// TIA Portal V17 export
FUNCTION_BLOCK "GraphTemplate"   // FB32000, GRAPH
VERSION : 0.1
// stored: AcknowledgeErrorsRequired true, AutoNumber false, GraphVersion 6.0, InitialValuesAcquisition false, IsIECCheckEnabled false, LanguageInNetworks LAD, LockOperatingMode false, PermanentILProcessingInMANMode false, SetENOAutomatically false, SkipSteps false, UDAEnableTagReadback false, WithAlarmHandling true
   // inherited from GRAPH_BASE
   VAR
      OFF_SQ_BASE : Bool;
   END_VAR
   VAR_INPUT
      OFF_SQ { ExternalWritable := 'False'} : Bool;
      INIT_SQ { ExternalWritable := 'False'} : Bool;
      ACK_EF { ExternalWritable := 'False'} : Bool;
      S_PREV { ExternalWritable := 'False'} : Bool;
      S_NEXT { ExternalWritable := 'False'} : Bool;
      SW_AUTO { ExternalWritable := 'False'} : Bool;
      SW_TAP { ExternalWritable := 'False'} : Bool;
      SW_TOP { ExternalWritable := 'False'} : Bool;
      SW_MAN { ExternalWritable := 'False'} : Bool;
      S_SEL { ExternalWritable := 'False'} : Int;
      S_ON { ExternalWritable := 'False'} : Bool;
      S_OFF { ExternalWritable := 'False'} : Bool;
      T_PUSH { ExternalWritable := 'False'} : Bool;
   END_VAR
   VAR_OUTPUT
      S_NO { ExternalWritable := 'False'} : Int;
      S_MORE { ExternalWritable := 'False'} : Bool;
      S_ACTIVE { ExternalWritable := 'False'} : Bool;
      ERR_FLT { ExternalWritable := 'False'} : Bool;
      AUTO_ON { ExternalWritable := 'False'} : Bool;
      TAP_ON { ExternalWritable := 'False'} : Bool;
      TOP_ON { ExternalWritable := 'False'} : Bool;
      MAN_ON { ExternalWritable := 'False'} : Bool;
   END_VAR
BEGIN
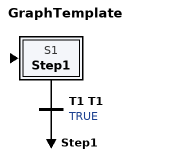
   // sequencer 1
   INITIAL_STEP Step1:   // S1
   END_STEP
   TRANSITION T1 FROM Step1 TO Step1   // T1
      := TRUE;
   END_TRANSITION
END_FUNCTION_BLOCK
